(* IEC 61131-3 sources: kns-pump-station/src/POUs/Station/FB_StationCore, 4 files *)

(* ---- FB_StationCore.decl.st ---- *)
// Назначение: ядро PRG_Station — порядок цикла станции (DESIGN, раздел 7, шаги 2–15) без обращений
//             к глобальным переменным: уставки (LKG с энергонезависимой копией, «Применить уставки
//             проекта», откат), команды станции и кнопки шкафа, режим, питание, защиты, действующее
//             управление, ступенчатое и ПИД (LIC101), чередование, АВР, задание частоты, блокировки,
//             вентиляция, тревоги KNS1.*, местная сигнализация, события журнала, состояние
//             stStationSts. Устройства — интерфейсами PL.I_MotorVfd и значениями входов, журнал —
//             I_StationEventSink, время — PL.I_TimeSource, данные GVL_Station и GVL_Persist —
//             параметрами VAR_IN_OUT: юнит-тесты идут с подменными насосами и временем, без модели и
//             сгенерированного слоя. Привязку к GVL_Devices, GVL_Hmi, GVL_IO, GVL_Persist, GVL_Log,
//             GVL_Sim, GVL_Time и GVL_DeviceList выполняет PRG_Station.
// Автор:      kr0nsch
// Версия:     0.3.0
// Документ:   docs/DESIGN.md, разделы 6.15 и 7; docs/04_algorithms.md, разделы 4, 15, 16, 18.3, 19
FUNCTION_BLOCK FB_StationCore
VAR_INPUT
    itfTime           : PL.I_TimeSource;      // GVL_Time.fbClockMain
    itfEvents         : I_StationEventSink;   // GVL_Log.fbEventLog
    aitfPump          : ARRAY[1..GVL_Const.STN_PUMP_COUNT] OF PL.I_MotorVfd;   // GVL_Devices.fbP101…fbP103
    axCommOk          : ARRAY[1..GVL_Const.STN_PUMP_COUNT] OF BOOL;   // нет MOT_WRN_COMM_LOSS в wWarning насоса
    axRunFeedback     : ARRAY[1..GVL_Const.STN_PUMP_COUNT] OF BOOL;   // GVL_IO.xP10n_RFB: подхват при старте ПЛК
    axPumpReset       : ARRAY[1..GVL_Const.STN_PUMP_COUNT] OF BOOL;   // GVL_Hmi.stP10nCmd.stCommon.xReset
    arCurrent_A       : ARRAY[1..GVL_Const.STN_PUMP_COUNT] OF REAL;   // fbIT1n1.rValue_eu
    axCurrentValid    : ARRAY[1..GVL_Const.STN_PUMP_COUNT] OF BOOL;   // fbIT1n1.xValid
    axOverheat        : ARRAY[1..GVL_Const.STN_PUMP_COUNT] OF BOOL;   // fbTS1n2.xValue
    rLevel_m          : REAL;                 // fbLT101.rValue_eu
    xLevelValid       : BOOL;                 // fbLT101.xValid
    eLevelNe107       : PL.E_Ne107Status;     // fbLT101.stSts.stCommon.eNe107
    xLevelL           : BOOL;                 // fbLT101.xL, xLL, xH, xHH
    xLevelLL          : BOOL;
    xLevelH           : BOOL;
    xLevelHH          : BOOL;
    rLvlL_m           : REAL;                 // GVL_Persist.stLT101Cfg: уставка L (порядок отметок)
    rLvlH_m           : REAL;                 // уставка H
    rLvlLProject_m    : REAL;                 // GVL_CfgProject.stLT101Cfg: уставка L проекта (цикл «Применить уставки
                                              // проекта»: LT101 восстанавливает PRG_Devices — после станции)
    rLvlHProject_m    : REAL;                 // уставка H проекта
    xFloatHigh        : BOOL;                 // fbLS102.xValue
    xFloatDry         : BOOL;                 // fbLS103.xValue
    xPowerOk          : BOOL;                 // fbES301.xValue
    xResetButton      : BOOL;                 // fbHS501.xValue (фронт выделяет ФБ)
    xSilenceButton    : BOOL;                 // fbHS502.xValue
    xGasHigh          : BOOL;                 // fbAT401.xH OR fbAT402.xH
    xDoorOpen         : BOOL;                 // fbZS404.xValue
    xTempHigh         : BOOL;                 // fbTT403.xH
    xFire             : BOOL;                 // fbYS405.xValue
    xApplyProjectCfg  : BOOL;                 // GVL_Hmi.xApplyProjectCfg (импульс сбрасывает PRG_Devices)
    xAckIdFound       : BOOL;                 // GVL_Log.fbAlarmSummary.AckById(stCmd.udiAckId) этого цикла
    xShelveIdFound    : BOOL;                 // … ShelveById(stCmd.udiShelveId, TRUE)
    xUnshelveIdFound  : BOOL;                 // … ShelveById(stCmd.udiUnshelveId, FALSE)
    xSimulation       : BOOL;                 // GVL_Sim.xSimulation
    udiSimFaultSeq    : UDINT;                // GVL_Sim.stSimSts.udiFaultSeq
    eLogExport        : E_LogExportState;     // GVL_Log.eExportState
    uiExportLines     : UINT;                 // GVL_Log.uiExportLines
    udiExportError    : UDINT;                // GVL_Log.udiExportError
    udiEventSeq       : UDINT;                // GVL_Log.fbEventLog.udiSeqLast
    udiLogOverwritten : UDINT;                // GVL_Log.fbEventLog.udiOverwritten
    auiUnack          : ARRAY[1..GVL_Const.ALM_PRIO_COUNT] OF UINT;   // GVL_Log.fbAlarmSummary (прошлый цикл)
    auiActive         : ARRAY[1..GVL_Const.ALM_PRIO_COUNT] OF UINT;
    ePrioUnack        : PL.E_AlarmPriority;
    udiNewHighSeq     : UDINT;
END_VAR
VAR_IN_OUT
    stCmd          : ST_StationCmd;           // GVL_Station.stStationCmd: импульсы и номера сбрасываются
    stCfgPersist   : ST_StationCfg;           // GVL_Persist.stStationCfg
    stCfgLkg       : ST_StationCfg;           // GVL_Station.stCfgLkg
    stCfgLkgRetain : ST_StationCfg;           // GVL_Persist.stStationCfgLkg: копия LKG, переживает перезапуск
    stRetain       : ST_StationRetain;        // GVL_Persist.stStationRetain
    fbLIC101       : PL.FB_PID;               // GVL_Station.fbLIC101
    stLIC101Cmd    : PL.ST_PidCmd;            // GVL_Station.stLIC101Cmd
    stLIC101Cfg    : PL.ST_PidCfg;            // GVL_Persist.stLIC101Cfg
    stLIC101Retain : PL.ST_DeviceRetain;      // GVL_Persist.stLIC101Retain
    fbAlarms       : FB_StationAlarms;        // GVL_Station.fbAlarms
END_VAR
VAR_OUTPUT
    stSts               : ST_StationSts;      // → GVL_Station.stStationSts
    axRun               : ARRAY[1..GVL_Const.STN_PUMP_COUNT] OF BOOL;   // → fbP10n.xAutoRun, GVL_Station.axPumpRun
    awInterlock         : ARRAY[1..GVL_Const.STN_PUMP_COUNT] OF WORD;   // → fbP10n.wInterlock, awPumpInterlock
    rSpeedSp_pct        : REAL;               // → fbP10n.rSpeedSpAuto_pct, GVL_Station.rSpeedSp_pct
    xSuppressFlowAlarms : BOOL;               // → fbPT201, fbFT202.xSuppressLimitAlarms
    xV1Run              : BOOL;               // → fbV1.xAutoRun
    wV1Interlock        : WORD;               // → fbV1.wInterlock
    xHorn               : BOOL;               // → GVL_IO.xHA1
    xLamp               : BOOL;               // → GVL_IO.xHL1
    xK1                 : BOOL;               // → GVL_IO.xK1 (TRUE — норма)
    xResetAllReq        : BOOL;               // импульс: Reset() всех GVL_DeviceList.aitfDevice
    xAckAllReq          : BOOL;               // импульс: AckAll() всех GVL_DeviceList.aitfDevice
    xExportReq          : BOOL;               // импульс: GVL_Log.fbEventLog.TakeSnapshot(), GVL_Log.xExportReq := TRUE
END_VAR
VAR
    fbMode         : FB_StationMode;          // 6.1
    fbPower        : FB_PowerRestore;         // 6.9
    fbProt         : FB_Protections;          // 6.7
    afbPumpProt    : ARRAY[1..GVL_Const.STN_PUMP_COUNT] OF FB_PumpProtection;   // 6.8
    fbSelect       : FB_ControlSelector;      // 6.2
    fbStepped      : FB_LevelControlStepped;  // 6.3
    fbPidCtl       : FB_LevelControlPid;      // 6.4
    fbRotation     : FB_PumpRotation;         // 6.5
    fbAts          : FB_Ats;                  // 6.6
    fbVent         : FB_Ventilation;          // 6.10
    fbAnnunciator  : FB_Annunciator;          // 6.12
    fbFlowSettle   : PL.FB_Delay;             // насос работает дольше STN_FLOW_SETTLE: давление и расход набраны
    xFirstCall     : BOOL := TRUE;            // первый вызов: старт приложения
    xResetBtnPrev  : BOOL;                    // HS501 прошлого вызова (фронт)
    xSilenceBtnPrev : BOOL;                   // HS502 прошлого вызова (фронт)
    uiRequiredPrev : UINT;                    // требуемое число прошлого цикла (FB_PowerRestore)
    eLogExportPrev : E_LogExportState;        // состояние выгрузки прошлого вызова (события 101019/101020)
    udiSimSeqPrev  : UDINT;                   // счётчик инъекций прошлого вызова (событие 101021)
    wCfgErr        : WORD;                    // ошибки уставок этого вызова
    eActPrev       : E_ControlAct;            // действующее управление прошлого вызова
END_VAR
VAR_TEMP
    uiPump         : UINT;                    // номер насоса
    uiCmdCount     : UINT;                    // обработано команд станции в этом вызове
    eCmdRes        : PL.E_CmdResult;          // результат последней команды
    xResetNow      : BOOL;                    // общий сброс в этом вызове (HS501 или HMI)
    xAckNow        : BOOL;                    // квитировать все (HMI)
    xSilenceNow    : BOOL;                    // «Звук» (HS502 или HMI)
    xCfgCmd        : BOOL;                    // уставки переписаны командой (событие уже записано)
    uiParam        : UINT;                    // номер изменённого параметра (событие 101017)
    rLvlLChk_m     : REAL;                    // L и H LT101 для проверки уставок станции (команда — уставки проекта)
    rLvlHChk_m     : REAL;
    wAckMask       : WORD;                    // маски команд тревог станции этого вызова
    wShelveMask    : WORD;
    wUnshelveMask  : WORD;
    uiRunningNow   : UINT;                    // работающие насосы
    axAdoptRun     : ARRAY[1..GVL_Const.STN_PUMP_COUNT] OF BOOL;   // «работает» для подхвата
    axTrip         : ARRAY[1..GVL_Const.STN_PUMP_COUNT] OF BOOL;   // фиксация недогрузки (KNS1.ULn)
    axAtsTrip      : ARRAY[1..GVL_Const.STN_PUMP_COUNT] OF BOOL;   // блокировка станции насоса (АВР)
    xAnyRunning    : BOOL;                    // работает хотя бы один насос
    xInitReq       : BOOL;                    // вход без рывка: смена управления или вход в «Автомат»
    xSteppedCont   : BOOL;                    // ступенчатый автомат продолжает работу (Restart <-> Stepped)
    eAct           : E_ControlAct;            // действующее управление
    uiRequired     : UINT;                    // требуемое число насосов
    uiTrack        : UINT;                    // «Ручной»: работающий насос с меньшей наработкой
    axCond         : ARRAY[1..GVL_Const.STN_ALARM_COUNT] OF BOOL;  // условия тревог KNS1.*
    axSuppress     : ARRAY[1..GVL_Const.STN_ALARM_COUNT] OF BOOL;  // подавления по условию
    arValue        : ARRAY[1..GVL_Const.STN_ALARM_COUNT] OF REAL;  // значения для событий
    uiSlot         : UINT;                    // слот тревоги
    xManual        : BOOL;                    // станция в «Ручном»
    eNe107         : PL.E_Ne107Status;        // сводный статус
    wState         : WORD;                    // биты STN_ST_*
    xMaint         : BOOL;                    // насосу нужно ТО
END_VAR

(* ---- ChangedParam.method.decl.st ---- *)
// Номер первого различающегося параметра уставок станции для события 101017 (04 §18.2: № 2–31 по
// порядку полей ST_StationCfg); таблица тревог или резерв — STN_CFG_PARAM_ALARMS; 0 — уставки
// совпадают. Сравнение по полям, без байтов выравнивания. Структуры — собственными параметрами
// метода (правило R2 контракта); метод без состояния, им пользуется и тест умолчаний
METHOD PUBLIC ChangedParam : UINT
VAR_IN_OUT CONSTANT
    stOld : ST_StationCfg;          // действующая копия
    stNew : ST_StationCfg;          // записанные уставки
END_VAR
VAR
    uiNo  : UINT;                   // номер параметра текущего поля
    uiIdx : UINT;                   // элемент массива
END_VAR

(* ---- ChangedParam.method.impl.st ---- *)
// Поля — по порядку раздела 18.2: номер растёт на 1 от поля к полю, первое отличие запоминается
ChangedParam := 0;
uiNo := GVL_Const.STN_CFG_PARAM_FIRST;
IF stNew.rLvlStop_m <> stOld.rLvlStop_m THEN
    ChangedParam := uiNo;                                           // № 2
END_IF
uiNo := uiNo + 1;
IF ChangedParam = 0 AND stNew.rLvlStartLead_m <> stOld.rLvlStartLead_m THEN
    ChangedParam := uiNo;
END_IF
uiNo := uiNo + 1;
IF ChangedParam = 0 AND stNew.rLvlStopAssist_m <> stOld.rLvlStopAssist_m THEN
    ChangedParam := uiNo;
END_IF
uiNo := uiNo + 1;
IF ChangedParam = 0 AND stNew.rLvlStartAssist_m <> stOld.rLvlStartAssist_m THEN
    ChangedParam := uiNo;
END_IF
uiNo := uiNo + 1;
IF ChangedParam = 0 AND stNew.tLvlConfirm <> stOld.tLvlConfirm THEN
    ChangedParam := uiNo;                                           // № 6
END_IF
uiNo := uiNo + 1;
IF ChangedParam = 0 AND stNew.rStepSpeed_pct <> stOld.rStepSpeed_pct THEN
    ChangedParam := uiNo;
END_IF
uiNo := uiNo + 1;
IF ChangedParam = 0 AND stNew.rLevelSp_m <> stOld.rLevelSp_m THEN
    ChangedParam := uiNo;                                           // № 8
END_IF
uiNo := uiNo + 1;
IF ChangedParam = 0 AND stNew.rAssistOn_pct <> stOld.rAssistOn_pct THEN
    ChangedParam := uiNo;
END_IF
uiNo := uiNo + 1;
IF ChangedParam = 0 AND stNew.tAssistOn <> stOld.tAssistOn THEN
    ChangedParam := uiNo;
END_IF
uiNo := uiNo + 1;
IF ChangedParam = 0 AND stNew.rAssistOff_pct <> stOld.rAssistOff_pct THEN
    ChangedParam := uiNo;
END_IF
uiNo := uiNo + 1;
IF ChangedParam = 0 AND stNew.tAssistOff <> stOld.tAssistOff THEN
    ChangedParam := uiNo;                                           // № 12
END_IF
uiNo := uiNo + 1;
IF ChangedParam = 0 AND stNew.uiDutyMax <> stOld.uiDutyMax THEN
    ChangedParam := uiNo;
END_IF
uiNo := uiNo + 1;
IF ChangedParam = 0 AND stNew.eRotation <> stOld.eRotation THEN
    ChangedParam := uiNo;
END_IF
uiNo := uiNo + 1;
IF ChangedParam = 0 AND stNew.tMaxContRun <> stOld.tMaxContRun THEN
    ChangedParam := uiNo;                                           // № 15
END_IF
uiNo := uiNo + 1;
IF ChangedParam = 0 AND stNew.tOverlap <> stOld.tOverlap THEN
    ChangedParam := uiNo;
END_IF
uiNo := uiNo + 1;
IF ChangedParam = 0 AND stNew.tStagger <> stOld.tStagger THEN
    ChangedParam := uiNo;
END_IF
uiNo := uiNo + 1;
IF ChangedParam = 0 AND stNew.tPwrRestart <> stOld.tPwrRestart THEN
    ChangedParam := uiNo;                                           // № 18
END_IF
uiNo := uiNo + 1;
IF ChangedParam = 0 AND stNew.tSeqStep <> stOld.tSeqStep THEN
    ChangedParam := uiNo;
END_IF
uiNo := uiNo + 1;
IF ChangedParam = 0 AND stNew.tPlcStart <> stOld.tPlcStart THEN
    ChangedParam := uiNo;
END_IF
uiNo := uiNo + 1;
IF ChangedParam = 0 AND stNew.tDryRelease <> stOld.tDryRelease THEN
    ChangedParam := uiNo;                                           // № 21
END_IF
uiNo := uiNo + 1;
IF ChangedParam = 0 AND stNew.rLdev102On_m <> stOld.rLdev102On_m THEN
    ChangedParam := uiNo;
END_IF
uiNo := uiNo + 1;
IF ChangedParam = 0 AND stNew.rLdev102Off_m <> stOld.rLdev102Off_m THEN
    ChangedParam := uiNo;
END_IF
uiNo := uiNo + 1;
IF ChangedParam = 0 AND stNew.rLdev103On_m <> stOld.rLdev103On_m THEN
    ChangedParam := uiNo;
END_IF
uiNo := uiNo + 1;
IF ChangedParam = 0 AND stNew.rLdev103Off_m <> stOld.rLdev103Off_m THEN
    ChangedParam := uiNo;                                           // № 25
END_IF
uiNo := uiNo + 1;
IF ChangedParam = 0 AND stNew.tLdev <> stOld.tLdev THEN
    ChangedParam := uiNo;
END_IF
uiNo := uiNo + 1;
IF ChangedParam = 0 AND stNew.tLtRecover <> stOld.tLtRecover THEN
    ChangedParam := uiNo;
END_IF
uiNo := uiNo + 1;
IF ChangedParam = 0 AND stNew.rUnderload_A <> stOld.rUnderload_A THEN
    ChangedParam := uiNo;                                           // № 28
END_IF
uiNo := uiNo + 1;
IF ChangedParam = 0 AND stNew.rUnderloadSpeed_pct <> stOld.rUnderloadSpeed_pct THEN
    ChangedParam := uiNo;
END_IF
uiNo := uiNo + 1;
IF ChangedParam = 0 AND stNew.tUnderload <> stOld.tUnderload THEN
    ChangedParam := uiNo;
END_IF
uiNo := uiNo + 1;
IF ChangedParam = 0 AND stNew.tV1Overrun <> stOld.tV1Overrun THEN
    ChangedParam := uiNo;                                           // № 31
END_IF

// Таблица тревог и резерв — один номер
IF ChangedParam = 0 THEN
    FOR uiIdx := 1 TO GVL_Const.STN_ALARM_COUNT DO
        IF stNew.astAlarm[uiIdx].ePriority <> stOld.astAlarm[uiIdx].ePriority
           OR stNew.astAlarm[uiIdx].tOnDelay <> stOld.astAlarm[uiIdx].tOnDelay
           OR stNew.astAlarm[uiIdx].tOffDelay <> stOld.astAlarm[uiIdx].tOffDelay
           OR stNew.astAlarm[uiIdx].tShelveMax <> stOld.astAlarm[uiIdx].tShelveMax THEN
            ChangedParam := GVL_Const.STN_CFG_PARAM_ALARMS;
        END_IF
    END_FOR
    FOR uiIdx := 0 TO GVL_Const.STN_CFG_RESERVE_REAL_LAST DO
        IF stNew.arReserve[uiIdx] <> stOld.arReserve[uiIdx] THEN
            ChangedParam := GVL_Const.STN_CFG_PARAM_ALARMS;
        END_IF
    END_FOR
    FOR uiIdx := 0 TO GVL_Const.STN_CFG_RESERVE_SHORT_LAST DO
        IF stNew.atReserve[uiIdx] <> stOld.atReserve[uiIdx] OR stNew.auiReserve[uiIdx] <> stOld.auiReserve[uiIdx] THEN
            ChangedParam := GVL_Const.STN_CFG_PARAM_ALARMS;
        END_IF
    END_FOR
END_IF

(* ---- FB_StationCore.impl.st ---- *)
// 0. Старт приложения (событие 101015) — первой записью станции
IF xFirstCall AND itfEvents <> 0 THEN
    itfEvents.LogEvent(eEvent := E_StationEvent.PlcStart, rValue := 0.0);
END_IF
uiCmdCount := 0;
eCmdRes := stSts.eCmdResult;

// 1. Уставки (DESIGN 7, шаг 2; 04 §18.3). «Применить уставки проекта» и откат командой переписывают
//    записанные уставки; корректные уставки становятся действующей копией (LKG), каждое принятое
//    изменение — событие 101017 (номер параметра; команда — значение 0). Копия LKG сохраняется в
//    энергонезависимой памяти (stCfgLkgRetain): при старте ПЛК действующая копия — сохранённая, если она
//    корректна, иначе уставки проекта; неверная правка, оставленная до перезапуска, не возвращает станцию
//    к уставкам проекта
IF xFirstCall THEN
    IF F_StationCfgCheck(stCfg := stCfgLkgRetain, stPidCfg := stLIC101Cfg, rLvlL_m := rLvlL_m,
                         rLvlH_m := rLvlH_m) = 0 THEN
        stCfgLkg := stCfgLkgRetain;
    ELSE
        stCfgLkg := GVL_StationDefaults.stStationCfg;
        stCfgLkgRetain := stCfgLkg;
    END_IF
END_IF
xCfgCmd := FALSE;
rLvlLChk_m := rLvlL_m;
rLvlHChk_m := rLvlH_m;
IF xApplyProjectCfg THEN
    stCfgPersist := GVL_StationDefaults.stStationCfg;
    stLIC101Cfg := GVL_StationDefaults.stLIC101Cfg;
    xCfgCmd := TRUE;
    // L/H LT101 уставок проекта восстанавливает PRG_Devices в этом же цикле, но после станции: уставки по умолчанию
    // проверяются по ним, а не по прежним (иначе ложная ошибка уставок на цикл и второе событие 101017)
    rLvlLChk_m := rLvlLProject_m;
    rLvlHChk_m := rLvlHProject_m;
END_IF
IF stCmd.xRevertCfg THEN
    stCfgPersist := stCfgLkg;
    uiCmdCount := uiCmdCount + 1;
    eCmdRes := PL.E_CmdResult.Accepted;
    xCfgCmd := TRUE;
    stCmd.xRevertCfg := FALSE;
END_IF
IF xCfgCmd AND itfEvents <> 0 THEN
    itfEvents.LogEvent(eEvent := E_StationEvent.CfgChanged, rValue := 0.0);
END_IF
wCfgErr := F_StationCfgCheck(stCfg := stCfgPersist, stPidCfg := stLIC101Cfg, rLvlL_m := rLvlLChk_m,
                             rLvlH_m := rLvlHChk_m);
IF wCfgErr = 0 THEN
    uiParam := ChangedParam(stOld := stCfgLkg, stNew := stCfgPersist);
    IF uiParam <> 0 THEN
        stCfgLkg := stCfgPersist;
        stCfgLkgRetain := stCfgPersist;                 // энергонезависимая копия — только при изменении
        // при старте записанные уставки принимаются молча; команда уже записала событие
        IF NOT xFirstCall AND NOT xCfgCmd AND itfEvents <> 0 THEN
            itfEvents.LogEvent(eEvent := E_StationEvent.CfgChanged, rValue := UINT_TO_REAL(uiParam));
        END_IF
    END_IF
END_IF

// 2. Команды станции и кнопки шкафа (DESIGN 7, шаг 3) — по порядку контракта 2.1: сброс,
//    квитирование, режим и способ, маски тревог, номера, звук, выгрузка
xResetNow := (xResetButton AND NOT xResetBtnPrev) OR stCmd.xResetAll;
IF xResetButton AND NOT xResetBtnPrev AND itfEvents <> 0 THEN
    itfEvents.LogEvent(eEvent := E_StationEvent.ResetAll, rValue := GVL_Const.STN_EVT_SRC_BUTTON);
END_IF
IF stCmd.xResetAll THEN
    uiCmdCount := uiCmdCount + 1;
    eCmdRes := PL.E_CmdResult.Accepted;
    IF itfEvents <> 0 THEN
        itfEvents.LogEvent(eEvent := E_StationEvent.ResetAll, rValue := GVL_Const.STN_EVT_SRC_HMI);
    END_IF
END_IF
IF xResetNow THEN
    fbLIC101.Reset();                                   // устройства — PRG_Station по xResetAllReq
END_IF
xResetAllReq := xResetNow;

xAckNow := stCmd.xAckAll;
IF xAckNow THEN
    uiCmdCount := uiCmdCount + 1;
    eCmdRes := PL.E_CmdResult.Accepted;
    fbLIC101.AckAll();
    IF itfEvents <> 0 THEN
        itfEvents.LogEvent(eEvent := E_StationEvent.AckAll, rValue := 0.0);
    END_IF
END_IF
xAckAllReq := xAckNow;

fbMode(xSetAuto := stCmd.xSetAuto, xSetManual := stCmd.xSetManual, xSetStepped := stCmd.xSetStepped,
       xSetLevelPid := stCmd.xSetLevelPid, aitfPump := aitfPump, itfEvents := itfEvents, stRetain := stRetain);
IF fbMode.uiCmdCount > 0 THEN
    uiCmdCount := uiCmdCount + fbMode.uiCmdCount;
    eCmdRes := fbMode.eCmdResult;
END_IF
xManual := fbMode.eMode <> E_StationMode.Auto;

wAckMask := stCmd.wAckReq;
wShelveMask := stCmd.wShelveReq;
wUnshelveMask := stCmd.wUnshelveReq;
IF wAckMask <> 0 THEN
    uiCmdCount := uiCmdCount + 1;
    eCmdRes := PL.E_CmdResult.Accepted;
END_IF
IF wShelveMask <> 0 THEN
    uiCmdCount := uiCmdCount + 1;
    eCmdRes := PL.E_CmdResult.Accepted;
END_IF
IF wUnshelveMask <> 0 THEN
    uiCmdCount := uiCmdCount + 1;
    eCmdRes := PL.E_CmdResult.Accepted;
END_IF

// номера тревог выполняет сводка (PRG_Station вызывает её до ядра): здесь — результат и сброс номера
IF stCmd.udiAckId <> 0 THEN
    uiCmdCount := uiCmdCount + 1;
    eCmdRes := SEL(xAckIdFound, PL.E_CmdResult.RejectedState, PL.E_CmdResult.Accepted);
END_IF
IF stCmd.udiShelveId <> 0 THEN
    uiCmdCount := uiCmdCount + 1;
    eCmdRes := SEL(xShelveIdFound, PL.E_CmdResult.RejectedState, PL.E_CmdResult.Accepted);
END_IF
IF stCmd.udiUnshelveId <> 0 THEN
    uiCmdCount := uiCmdCount + 1;
    eCmdRes := SEL(xUnshelveIdFound, PL.E_CmdResult.RejectedState, PL.E_CmdResult.Accepted);
END_IF

xSilenceNow := (xSilenceButton AND NOT xSilenceBtnPrev) OR stCmd.xSilence;
IF xSilenceButton AND NOT xSilenceBtnPrev AND itfEvents <> 0 THEN
    itfEvents.LogEvent(eEvent := E_StationEvent.Silence, rValue := GVL_Const.STN_EVT_SRC_BUTTON);
END_IF
IF stCmd.xSilence THEN
    uiCmdCount := uiCmdCount + 1;
    eCmdRes := PL.E_CmdResult.Accepted;
    IF itfEvents <> 0 THEN
        itfEvents.LogEvent(eEvent := E_StationEvent.Silence, rValue := GVL_Const.STN_EVT_SRC_HMI);
    END_IF
END_IF

// выгрузка журнала: пока идёт прежняя (снимок или запись), новая отклоняется
xExportReq := FALSE;
IF stCmd.xExportLog THEN
    uiCmdCount := uiCmdCount + 1;
    IF eLogExport = E_LogExportState.Snapshot OR eLogExport = E_LogExportState.Writing THEN
        eCmdRes := PL.E_CmdResult.RejectedState;
    ELSE
        eCmdRes := PL.E_CmdResult.Accepted;
        xExportReq := TRUE;
    END_IF
END_IF

// импульсы и номера сброшены в том же цикле (04 §19.2)
stCmd.xSetAuto := FALSE;
stCmd.xSetManual := FALSE;
stCmd.xSetStepped := FALSE;
stCmd.xSetLevelPid := FALSE;
stCmd.xAckAll := FALSE;
stCmd.xResetAll := FALSE;
stCmd.xSilence := FALSE;
stCmd.xExportLog := FALSE;
stCmd.wAckReq := 0;
stCmd.wShelveReq := 0;
stCmd.wUnshelveReq := 0;
stCmd.udiAckId := 0;
stCmd.udiShelveId := 0;
stCmd.udiUnshelveId := 0;
xResetBtnPrev := xResetButton;
xSilenceBtnPrev := xSilenceButton;

// 3. Насосы: работающие (в первом вызове устройства ещё не вызывались — по ОС GVL_IO.xP10n_RFB)
uiRunningNow := 0;
xAnyRunning := FALSE;
FOR uiPump := 1 TO GVL_Const.STN_PUMP_COUNT DO
    axAdoptRun[uiPump] := axRunFeedback[uiPump];
    IF NOT xFirstCall THEN
        axAdoptRun[uiPump] := FALSE;
        IF aitfPump[uiPump] <> 0 THEN
            axAdoptRun[uiPump] := aitfPump[uiPump].Running;
        END_IF
    END_IF
    IF axAdoptRun[uiPump] THEN
        uiRunningNow := uiRunningNow + 1;
        xAnyRunning := TRUE;
    END_IF
END_FOR

// 4. Питание (требуемое число — прошлого цикла), защиты, защиты насосов (DESIGN 7, шаг 5)
fbPower(xPowerOk := xPowerOk, uiRequired := uiRequiredPrev, uiRunningRequested := fbRotation.uiRunningRequested,
        itfTime := itfTime, itfEvents := itfEvents, stCfg := stCfgLkg);
fbProt(rLevel_m := rLevel_m, xLevelValid := xLevelValid, eLevelNe107 := eLevelNe107, xLevelL := xLevelL,
       xLevelLL := xLevelLL, xLevelH := xLevelH, xLevelHH := xLevelHH, xFloatHigh := xFloatHigh,
       xFloatDry := xFloatDry, uiRunning := uiRunningNow, itfTime := itfTime, itfEvents := itfEvents,
       stCfg := stCfgLkg);
FOR uiPump := 1 TO GVL_Const.STN_PUMP_COUNT DO
    IF aitfPump[uiPump] <> 0 THEN
        afbPumpProt[uiPump](xRunning := aitfPump[uiPump].Running, rSpeedAct_pct := aitfPump[uiPump].SpeedAct,
                            rCurrent_A := arCurrent_A[uiPump], xCurrentValid := axCurrentValid[uiPump],
                            xOverheat := axOverheat[uiPump], xReset := axPumpReset[uiPump] OR xResetNow,
                            itfTime := itfTime, stCfg := stCfgLkg);
    ELSE
        afbPumpProt[uiPump](xRunning := FALSE, rSpeedAct_pct := 0.0, rCurrent_A := arCurrent_A[uiPump],
                            xCurrentValid := FALSE, xOverheat := axOverheat[uiPump],
                            xReset := axPumpReset[uiPump] OR xResetNow, itfTime := itfTime, stCfg := stCfgLkg);
    END_IF
    axTrip[uiPump] := afbPumpProt[uiPump].xUnderloadTrip;
    // АВР — по отказу устройства или блокировке станции насоса: недогрузка и перегрев. TS1n2 без задержки приходит
    // раньше аварии ПЧ (фильтр tExtFaultFilter): насос останавливается и теряет запрос до отказа (04 §9.1, PMI-16)
    axAtsTrip[uiPump] := afbPumpProt[uiPump].wInterlock <> 0;
END_FOR

// 5. Действующее управление (готовность ПИД — прошлого цикла); смена управления или вход в
//    «Автомат» — вход без рывка: число насосов по работающим, роли — работающим (шаг 6)
fbSelect(eMode := fbMode.eMode, eMethod := fbMode.eMethod, xPowerLost := fbPower.xPowerLost,
         xRestart := fbPower.xRestart, xDryRun := fbProt.xDryRun, xFloatMode := fbProt.xFloatMode,
         xEmergency := fbProt.xEmergency, xPidReady := fbPidCtl.xPidReady);
eAct := fbSelect.eControlAct;
xInitReq := fbSelect.xChanged OR fbMode.xEnteredAuto;
// последовательный пуск идёт по тому же ступенчатому автомату: Restart <-> Stepped — без новой инициализации
xSteppedCont := (eAct = E_ControlAct.Stepped OR eAct = E_ControlAct.Restart)
                AND (eActPrev = E_ControlAct.Stepped OR eActPrev = E_ControlAct.Restart);

// 6. Регуляторы вызываются всегда (таймеры непрерывны); уровень — годный по защитам (LT101 не
//    исключён). Последовательный пуск — по ступенчатому автомату: ПИД в слежении (шаг 7)
fbStepped(xEnable := eAct = E_ControlAct.Stepped OR eAct = E_ControlAct.Restart, rLevel_m := rLevel_m,
          xLevelValid := fbProt.xLevelUsable, xInit := xInitReq AND NOT xSteppedCont, uiInitPumps := uiRunningNow,
          itfTime := itfTime, stCfg := stCfgLkg);
fbPidCtl(xEnable := eAct = E_ControlAct.LevelPid, rLevel_m := rLevel_m, xLevelValid := fbProt.xLevelUsable,
         rPidOut_pct := fbLIC101.rOut_pct, ePidMode := fbLIC101.Mode, aitfPump := aitfPump, axCommOk := axCommOk,
         uiLead := fbRotation.uiLead, xInit := xInitReq, uiInitPumps := uiRunningNow,
         xPowerRestore := fbPower.xPowerLost OR fbPower.xRestart, itfTime := itfTime, stCfg := stCfgLkg);
CASE eAct OF
    E_ControlAct.Stepped:
        uiRequired := fbStepped.uiRequired;
    E_ControlAct.Restart:
        // последовательный пуск охватывает все насосы состояния под ним: сухой ход — 0, по поплавкам и аварийный
        // уровень — все (ведущий, подпорный, остальные), иначе ступенчатый автомат; по одному — uiRequestLimit
        IF fbProt.xDryRun THEN
            uiRequired := 0;
        ELSIF fbProt.xFloatMode THEN
            uiRequired := fbProt.uiFloatRequired;
        ELSIF fbProt.xEmergency THEN
            uiRequired := GVL_Const.STN_PUMP_COUNT;
        ELSE
            uiRequired := fbStepped.uiRequired;
        END_IF
    E_ControlAct.LevelPid:
        uiRequired := fbPidCtl.uiRequired;
    E_ControlAct.Emergency:
        uiRequired := GVL_Const.STN_PUMP_COUNT;
    E_ControlAct.Float:
        uiRequired := fbProt.uiFloatRequired;
ELSE
    uiRequired := 0;                                    // DryRunStop, PowerLost, Manual
END_CASE

// 7. Роли и чередование (шаг 8): старт ПЛК — подхват по ОС; АВР (шаг 9)
fbRotation(xEnable := NOT xManual, uiRequired := uiRequired, uiRequestLimit := fbPower.uiRequestLimit,
           xRequireComm := eAct = E_ControlAct.LevelPid,
           xHandoverAllowed := eAct = E_ControlAct.Stepped OR eAct = E_ControlAct.LevelPid,
           xAdopt := xInitReq OR xFirstCall, axAdoptRun := axAdoptRun, aitfPump := aitfPump, axCommOk := axCommOk,
           itfTime := itfTime, itfEvents := itfEvents, stCfg := stCfgLkg, stRetain := stRetain);
fbAts(xEnable := NOT xManual, aitfPump := aitfPump, axRun := fbRotation.axRun, axTrip := axAtsTrip,
      uiRequired := uiRequired, uiAvailable := fbRotation.uiAvailable, uiForeign := fbRotation.uiForeign,
      itfTime := itfTime, itfEvents := itfEvents, stCfg := stCfgLkg);

// 8. LIC101 (шаг 10; 04 §7.1): задание — внешнее из LKG, слежение за ведущим, когда ПИД не управляет
fbLIC101(rPv_eu := rLevel_m, xPvValid := fbProt.xLevelUsable, xSpExt := TRUE, rSpExt_eu := stCfgLkg.rLevelSp_m,
         xTrack := fbPidCtl.xTrack, rTrack_pct := fbPidCtl.rTrack_pct, rOutAct_pct := fbPidCtl.rTrack_pct,
         itfTime := itfTime, stCmd := stLIC101Cmd, stCfg := stLIC101Cfg, stRetain := stLIC101Retain);

// 9. Общее задание частоты (шаг 11). «Ручной» — задание работающего насоса с меньшей наработкой
//    (будущего ведущего): вход в «Автомат» без рывка (04 §3.2); сухой ход и нет напряжения — прежнее
CASE eAct OF
    E_ControlAct.LevelPid:
        rSpeedSp_pct := fbLIC101.rOut_pct;
    E_ControlAct.Stepped:
        rSpeedSp_pct := stCfgLkg.rStepSpeed_pct;
    E_ControlAct.Restart:
        // последовательный пуск при аварийном уровне или по поплавкам — на полной частоте, как сами эти режимы
        IF (fbProt.xFloatMode OR fbProt.xEmergency) AND NOT fbProt.xDryRun THEN
            rSpeedSp_pct := GVL_Const.STN_FULL_SPEED_PCT;
        ELSE
            rSpeedSp_pct := stCfgLkg.rStepSpeed_pct;
        END_IF
    E_ControlAct.Emergency, E_ControlAct.Float:
        rSpeedSp_pct := GVL_Const.STN_FULL_SPEED_PCT;
    E_ControlAct.Manual:
        uiTrack := 0;
        FOR uiPump := 1 TO GVL_Const.STN_PUMP_COUNT DO
            IF aitfPump[uiPump] <> 0 THEN
                IF aitfPump[uiPump].Running THEN
                    IF uiTrack = 0 THEN
                        uiTrack := uiPump;
                    ELSIF aitfPump[uiPump].RunSeconds < aitfPump[uiTrack].RunSeconds THEN
                        uiTrack := uiPump;
                    END_IF
                END_IF
            END_IF
        END_FOR
        IF uiTrack <> 0 THEN
            rSpeedSp_pct := aitfPump[uiTrack].SpeedRef;
        END_IF
ELSE
    ;                                                   // DryRunStop, PowerLost: запросов нет
END_CASE

// 10. Входы автоматики устройств (шаг 12): запросы, блокировки, подавление тревог коллектора, В1
FOR uiPump := 1 TO GVL_Const.STN_PUMP_COUNT DO
    axRun[uiPump] := fbRotation.axRun[uiPump];
    awInterlock[uiPump] := afbPumpProt[uiPump].wInterlock;
    IF fbProt.xDryRun THEN
        awInterlock[uiPump] := awInterlock[uiPump] OR GVL_Const.KNS_ILK_DRY_RUN;
    END_IF
END_FOR
fbFlowSettle(xIn := xAnyRunning, tOnDelay := GVL_Const.STN_FLOW_SETTLE, itfTime := itfTime);
xSuppressFlowAlarms := NOT fbFlowSettle.xOut;
fbVent(xGasHigh := xGasHigh, xDoorOpen := xDoorOpen, xTempHigh := xTempHigh, xFire := xFire, itfTime := itfTime,
       stCfg := stCfgLkg);
xV1Run := fbVent.xRun;
wV1Interlock := fbVent.wInterlock;

// 11. Тревоги KNS1.* (шаг 13; условия и подавления — 04 §15, DESIGN 6.11)
FOR uiSlot := 1 TO GVL_Const.STN_ALARM_COUNT DO
    axCond[uiSlot] := FALSE;
    axSuppress[uiSlot] := FALSE;
    arValue[uiSlot] := 0.0;
END_FOR
// режим по поплавкам — управление только в «Автомате»: там срабатывания поплавков — штатные точки управления; в
// «Ручном» автоматика по поплавкам насосы не пускает, EHL (Critical) и DRY нужны оператору (04 §3.1, §10.2)
axCond[E_StationAlarm.EHL] := fbProt.xEmergency;
axSuppress[E_StationAlarm.EHL] := fbProt.xFloatMode AND NOT xManual;
arValue[E_StationAlarm.EHL] := rLevel_m;
axCond[E_StationAlarm.DRY] := fbProt.xDryRun;
axSuppress[E_StationAlarm.DRY] := fbProt.xFloatMode AND NOT xManual;
arValue[E_StationAlarm.DRY] := rLevel_m;
axCond[E_StationAlarm.LACK] := fbAts.xLack;
axSuppress[E_StationAlarm.LACK] := fbPower.xPowerLost OR xManual;
arValue[E_StationAlarm.LACK] := UINT_TO_REAL(uiRequired);
axCond[E_StationAlarm.NORES] := fbAts.xNoReserve;
// сухой ход станции блокирует все насосы: они недоступны по защите, а не из-за отказов (дубль KNS1.DRY)
axSuppress[E_StationAlarm.NORES] := fbAts.xLack OR fbPower.xPowerLost OR xManual OR fbProt.xDryRun;
arValue[E_StationAlarm.NORES] := UINT_TO_REAL(fbRotation.uiAvailable);
axCond[E_StationAlarm.ATS] := fbAts.xAtsActive;
axSuppress[E_StationAlarm.ATS] := fbPower.xPowerLost;
arValue[E_StationAlarm.ATS] := UDINT_TO_REAL(fbAts.udiAtsCount);
axCond[E_StationAlarm.FLOAT] := fbProt.xFloatMode;
axCond[E_StationAlarm.LDEV] := fbProt.xLdev;
arValue[E_StationAlarm.LDEV] := WORD_TO_REAL(fbProt.wLdev);
axCond[E_StationAlarm.STEP] := fbSelect.xStepFallback;
// последовательный пуск идёт по ступенчатому автомату при любой готовности ПИД (04 §4) — не деградация
axSuppress[E_StationAlarm.STEP] := eAct = E_ControlAct.Emergency OR eAct = E_ControlAct.Float
                                   OR eAct = E_ControlAct.DryRunStop OR eAct = E_ControlAct.PowerLost
                                   OR eAct = E_ControlAct.Restart;
axCond[E_StationAlarm.NOAUTO] := xManual;
FOR uiPump := 1 TO GVL_Const.STN_PUMP_COUNT DO
    axCond[E_StationAlarm.UL1 + uiPump - 1] := axTrip[uiPump];
    arValue[E_StationAlarm.UL1 + uiPump - 1] := arCurrent_A[uiPump];
END_FOR
axCond[E_StationAlarm.SIM] := xSimulation;
fbAlarms(axCond := axCond, axSuppress := axSuppress, arValue := arValue, wAckReq := wAckMask,
         wShelveReq := wShelveMask, wUnshelveReq := wUnshelveMask, xAckAll := xAckNow OR xResetNow,
         itfTime := itfTime, stCfg := stCfgLkg);
fbAnnunciator(auiUnack := auiUnack, auiActive := auiActive, udiNewHighSeq := udiNewHighSeq,
              xSilence := xSilenceNow, itfTime := itfTime);
xHorn := fbAnnunciator.xHorn;
xLamp := fbAnnunciator.xLamp;
xK1 := fbAnnunciator.xK1Energized;

// 12. События журнала (шаг 14): выгрузка CSV завершена или с ошибкой; изменена инъекция отказа
IF eLogExport <> eLogExportPrev AND itfEvents <> 0 THEN
    IF eLogExport = E_LogExportState.Done THEN
        itfEvents.LogEvent(eEvent := E_StationEvent.LogExported, rValue := UINT_TO_REAL(uiExportLines));
    ELSIF eLogExport = E_LogExportState.Error THEN
        itfEvents.LogEvent(eEvent := E_StationEvent.LogExportFailed, rValue := UDINT_TO_REAL(udiExportError));
    END_IF
END_IF
eLogExportPrev := eLogExport;
IF NOT xFirstCall AND udiSimFaultSeq <> udiSimSeqPrev AND itfEvents <> 0 THEN
    itfEvents.LogEvent(eEvent := E_StationEvent.SimFaultChanged, rValue := UDINT_TO_REAL(udiSimFaultSeq));
END_IF
udiSimSeqPrev := udiSimFaultSeq;

// 13. Состояние станции (шаг 15; 04 §19.3)
wState := 0;
IF fbProt.xDryRun THEN
    wState := wState OR GVL_Const.STN_ST_DRY_RUN;
END_IF
IF fbProt.xEmergency THEN
    wState := wState OR GVL_Const.STN_ST_EMERGENCY;
END_IF
IF fbProt.xFloatMode THEN
    wState := wState OR GVL_Const.STN_ST_FLOAT;
END_IF
IF axCond[E_StationAlarm.STEP] AND NOT axSuppress[E_StationAlarm.STEP] THEN
    wState := wState OR GVL_Const.STN_ST_STEP_FALLBACK;
END_IF
IF fbPower.xPowerLost THEN
    wState := wState OR GVL_Const.STN_ST_POWER_LOST;
END_IF
IF fbPower.xRestart THEN
    wState := wState OR GVL_Const.STN_ST_RESTART;
END_IF
IF fbAts.xAtsActive THEN
    wState := wState OR GVL_Const.STN_ST_ATS;
END_IF
IF axCond[E_StationAlarm.NORES] AND NOT axSuppress[E_StationAlarm.NORES] THEN
    wState := wState OR GVL_Const.STN_ST_NO_RESERVE;
END_IF
IF axCond[E_StationAlarm.LACK] AND NOT axSuppress[E_StationAlarm.LACK] THEN
    wState := wState OR GVL_Const.STN_ST_LACK;
END_IF
IF fbProt.xLs102Masked THEN
    wState := wState OR GVL_Const.STN_ST_LS102_MASKED;
END_IF
IF fbProt.xLs103Masked THEN
    wState := wState OR GVL_Const.STN_ST_LS103_MASKED;
END_IF
IF xSimulation THEN
    wState := wState OR GVL_Const.STN_ST_SIMULATION;
END_IF
IF xHorn THEN
    wState := wState OR GVL_Const.STN_ST_HORN;
END_IF
IF NOT xK1 THEN
    wState := wState OR GVL_Const.STN_ST_COMMON_ALARM;
END_IF
IF ePrioUnack <> PL.E_AlarmPriority.None THEN
    wState := wState OR GVL_Const.STN_ST_UNACK;
END_IF

// NE 107 станции: F — LACK; C — «Ручной», имитация, ошибка уставок; S — FLOAT, STEP, LDEV, NORES;
// M — ТО насоса. Тревога учитывается после своей задержки и без подавления по условию
eNe107 := PL.E_Ne107Status.Good;
xMaint := FALSE;
FOR uiPump := 1 TO GVL_Const.STN_PUMP_COUNT DO
    IF aitfPump[uiPump] <> 0 THEN
        xMaint := xMaint OR aitfPump[uiPump].Status = PL.E_Ne107Status.MaintenanceRequired;
    END_IF
END_FOR
IF xMaint THEN
    eNe107 := PL.E_Ne107Status.MaintenanceRequired;
END_IF
IF ((fbAlarms.wAlmActive AND SHL(WORD#1, E_StationAlarm.FLOAT - 1)) <> 0 AND NOT axSuppress[E_StationAlarm.FLOAT])
   OR ((fbAlarms.wAlmActive AND SHL(WORD#1, E_StationAlarm.STEP - 1)) <> 0 AND NOT axSuppress[E_StationAlarm.STEP])
   OR ((fbAlarms.wAlmActive AND SHL(WORD#1, E_StationAlarm.LDEV - 1)) <> 0 AND NOT axSuppress[E_StationAlarm.LDEV])
   OR ((fbAlarms.wAlmActive AND SHL(WORD#1, E_StationAlarm.NORES - 1)) <> 0
       AND NOT axSuppress[E_StationAlarm.NORES]) THEN
    eNe107 := PL.F_Ne107Worst(eA := eNe107, eB := PL.E_Ne107Status.OutOfSpecification);
END_IF
IF xManual OR xSimulation OR wCfgErr <> 0 THEN
    eNe107 := PL.F_Ne107Worst(eA := eNe107, eB := PL.E_Ne107Status.CheckFunction);
END_IF
IF (fbAlarms.wAlmActive AND SHL(WORD#1, E_StationAlarm.LACK - 1)) <> 0 AND NOT axSuppress[E_StationAlarm.LACK] THEN
    eNe107 := PL.E_Ne107Status.Failure;
END_IF

stSts.eMode := fbMode.eMode;
stSts.eMethod := fbMode.eMethod;
stSts.eControlAct := eAct;
stSts.eNe107 := eNe107;
stSts.wState := wState;
stSts.wCfgErr := wCfgErr;
FOR uiPump := 1 TO GVL_Const.STN_PUMP_COUNT DO
    stSts.aeRole[uiPump] := fbRotation.aeRole[uiPump];
END_FOR
stSts.uiPumpsRequired := uiRequired;
stSts.uiPumpsRunning := fbRotation.uiRunning;
stSts.uiPumpsAvailable := fbRotation.uiAvailable;
stSts.uiLeadPump := fbRotation.uiLead;
stSts.uiSeqRemain_s := fbPower.uiSeqRemain_s;
stSts.eCmdResult := eCmdRes;
stSts.uiCmdSeq := stSts.uiCmdSeq + uiCmdCount;     // UINT по кругу (контракт 2.1)
stSts.wAlmActive := fbAlarms.wAlmActive;
stSts.wAlmUnack := fbAlarms.wAlmUnack;
stSts.wAlmShelved := fbAlarms.wAlmShelved;
stSts.ePrioUnack := ePrioUnack;
FOR uiSlot := 1 TO GVL_Const.ALM_PRIO_COUNT DO
    stSts.auiUnack[uiSlot] := auiUnack[uiSlot];
END_FOR
stSts.eLogExport := eLogExport;
stSts.rLevel_m := rLevel_m;
stSts.rLevelSp_m := stCfgLkg.rLevelSp_m;
stSts.rSpeedSp_pct := rSpeedSp_pct;
stSts.udiEventSeq := udiEventSeq;
stSts.udiLogOverwritten := udiLogOverwritten;

uiRequiredPrev := uiRequired;
eActPrev := eAct;
xFirstCall := FALSE;
